// TIA Portal V20 export
// export: Created 2026-10-20T12:44:28.6307015Z, ExportSetting WithDefaults, DisplayName Totally Integrated Automation Portal, DisplayVersion V20 Update 6, DisplayName TIA Portal Openness, DisplayVersion V20 Update 6, DisplayName TIA Portal Version Control Interface, DisplayVersion V20 Update 6, DisplayName SINAMICS Startdrive Advanced, DisplayVersion V20 SP1, DisplayName SINAMICS Startdrive G130, G150, S120, S150, SINAMICS MV, G220, S200, S210, DisplayVersion V20 SP1, DisplayName SINAMICS Startdrive G110M, G120, G120C, G120D, G120P, G115D, DisplayVersion V20 SP1, DisplayName STEP 7 Professional, DisplayVersion V20 Update 6, DisplayName STEP 7 Safety, DisplayVersion V20 Update 2, DisplayName WinCC Basic/Comfort/Advanced, DisplayVersion V20 Update 6, DisplayName WinCC Unified, DisplayVersion V20 Update 6
FUNCTION "Set_Bit_F" : Void   // FC7, SCL
{ S7_Optimized_Access := 'TRUE' }
VERSION : 0.1
// stored: AutoNumber true, IsIECCheckEnabled false, SetENOAutomatically false, UDAEnableTagReadback false
   VAR_INPUT
      Bit : UInt;
      Bit_Value : Bool;
   END_VAR
   VAR_IN_OUT
      Var : Word;
   END_VAR
BEGIN
   IF #Bit_Value THEN
       // Set the bit
       #Var := #Var OR SHL(IN := WORD#1, N := #Bit);
   // ELSE
   //     // Reset the bit
   //     #Var := #Var OR SHL(IN := DWORD#1, N := #Bit);
   END_IF;
END_FUNCTION
